// TIA Portal V21 export
// export: Created 2026-11-07T17:04:58.6788832Z, ExportSetting WithDefaults, DisplayName Totally Integrated Automation Portal, DisplayVersion V21, DisplayName STEP 7 Professional, DisplayVersion V21, DisplayName STEP 7 Safety, DisplayVersion V21, DisplayName Tech WebApplication, DisplayVersion V21, DisplayName WinCC Basic/Comfort/Advanced, DisplayVersion V21, DisplayName WinCC Unified, DisplayVersion V21
TextList "TL_BalMode"  ListRange=Decimal
  TextListEntry   EntryType=SingleValue, Text="0 lijevo/desno"
  TextListEntry   EntryType=SingleValue, From=1, To=1, Text="1 + pramac/krma"
